(*~
	<docu>
		<summary>
			Reset command (command bit 0). Never blocked; aborts any other running command.
		</summary>
	</docu>
~*)
FUNCTION_BLOCK TcoAteqG6_ResetTask_v_3_5_x EXTENDS TcoAteqG6Task_v_3_5_x

IF Execute() THEN
	IF CheckReferences() THEN
		// AX step 0: reset handshake
		IF _progress = 0 THEN
			inoStatus.ActionDescription := '<#Resetting instrument#>';
			IF Handshake(MASK_RESET) THEN
				GoTo(100);
			END_IF
		END_IF

		// AX step 100
		IF _progress = 100 THEN
			inoStatus.ActionDescription := '<#Instrument reset#>';
			DoneWhen(TRUE);
		END_IF
		Supervise();
	END_IF
END_IF

IF THIS^.Error AND NOT _errorMessage.Pinned THEN
	THIS^.Restore();
END_IF

METHOD FB_init : BOOL
VAR_INPUT
	bInitRetains : BOOL; // if TRUE, the retain variables are initialized (warm start / cold start)
	bInCopyCode : BOOL;  // if TRUE, the instance afterwards gets moved into the copy code (online change)
	ParentObject : ITcoObject;
END_VAR
END_METHOD

END_FUNCTION_BLOCK

(* stored: Version 1.1.0.1, ProductVersion 3.1.4024.12
   POU TcoAteqG6_ResetTask_v_3_5_x: Id {22df437c-dc0b-4448-9ce5-135934773db5}, SpecialFunc None
   Method FB_init: Id {ed9cb579-8066-48ab-980b-330a1f5972e6} *)
